Fanuc KAREL source: kx00016.KL

-- PROVISIONAL review KL for V770-1; original PC SHA256 9ae1134a2e4d204c49ba62ba8c96c66653911a0fe4342274def18d15bde58f1a
-- Incomplete behavior may be omitted. Consult companion uncertainty JSON. Do not deploy.
PROGRAM KX00016
%NOLOCKGROUP
VAR
  I : INTEGER
  J : INTEGER
  B : BOOLEAN
  F : FILE
  S : STRING[80]
-- UNRESOLVED_DECL P type=000102
BEGIN
  -- UNRESOLVED_PC offsets 5-7; opcodes 9D,0D
  -- UNRESOLVED_PC offsets 12-16; opcodes 7F
END KX00016
